FUNCTION_BLOCK Model (* Composite Function Block Type *)
  (* Standard: 61499-2 *)
  (* Version 0.0, 7/13/2016, Andrei, nxtControl GmbH, template *)
  PACKAGE Main;
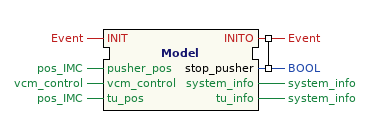
  EVENT_INPUT
    INIT; (* Initialization Request *)
  END_EVENT
  EVENT_OUTPUT
    INITO WITH stop_pusher; (* Initialization Confirm *)
  END_EVENT
  VAR_OUTPUT
    stop_pusher : BOOL;
  END_VAR
  SOCKETS
    pusher_pos : pos_IMC;
    vcm_control : vcm_control;
    tu_pos : pos_IMC;
  END_SOCKETS
  PLUGS
    system_info : system_info;
    tu_info : system_info;
  END_PLUGS
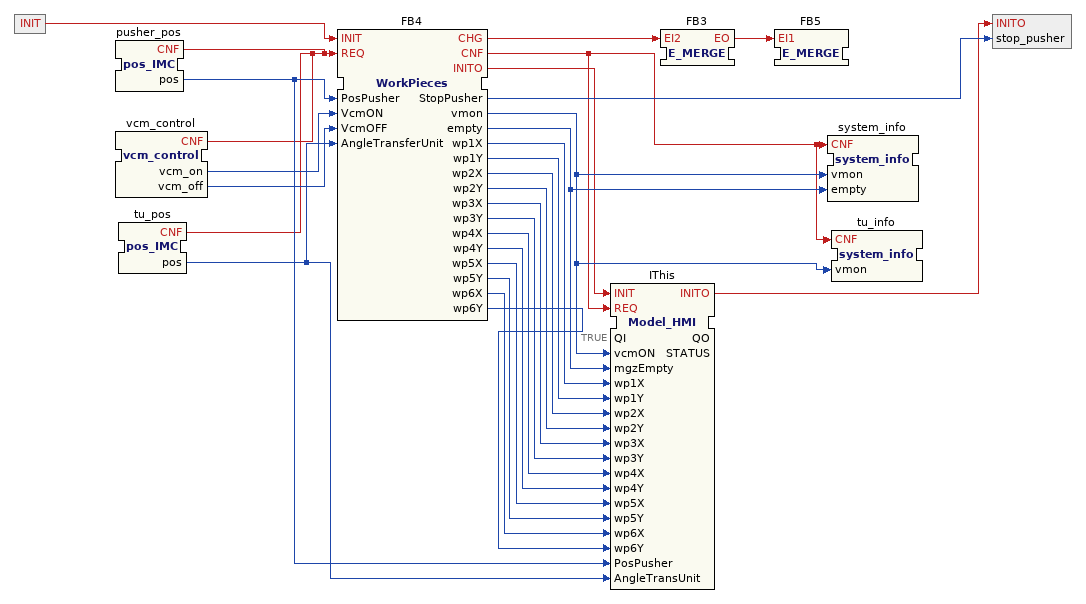
  FBS
    FB3 : E_MERGE;
    FB5 : E_MERGE;
    FB4 : WorkPieces;
    IThis : Model_HMI(QI := TRUE);
  END_FBS
  EVENT_CONNECTIONS
    FB4.CHG TO FB3.EI2;
    FB3.EO TO FB5.EI1;
    INIT TO FB4.INIT;
    pusher_pos.CNF TO FB4.REQ;
    vcm_control.CNF TO FB4.REQ;
    tu_pos.CNF TO FB4.REQ;
    FB4.CNF TO system_info.CNF;
    FB4.INITO TO IThis.INIT;
    FB4.CNF TO IThis.REQ;
    IThis.INITO TO INITO;
    FB4.CNF TO tu_info.CNF;
  END_CONNECTIONS
  DATA_CONNECTIONS
    FB4.StopPusher TO stop_pusher;
    pusher_pos.pos TO FB4.PosPusher;
    vcm_control.vcm_on TO FB4.VcmON;
    vcm_control.vcm_off TO FB4.VcmOFF;
    tu_pos.pos TO FB4.AngleTransferUnit;
    FB4.vmon TO system_info.vmon;
    FB4.empty TO system_info.empty;
    FB4.vmon TO IThis.vcmON;
    FB4.empty TO IThis.mgzEmpty;
    FB4.wp1X TO IThis.wp1X;
    FB4.wp1Y TO IThis.wp1Y;
    FB4.wp2X TO IThis.wp2X;
    FB4.wp2Y TO IThis.wp2Y;
    FB4.wp3X TO IThis.wp3X;
    FB4.wp3Y TO IThis.wp3Y;
    FB4.wp4X TO IThis.wp4X;
    FB4.wp4Y TO IThis.wp4Y;
    FB4.wp5X TO IThis.wp5X;
    FB4.wp5Y TO IThis.wp5Y;
    FB4.wp6X TO IThis.wp6X;
    FB4.wp6Y TO IThis.wp6Y;
    pusher_pos.pos TO IThis.PosPusher;
    tu_pos.pos TO IThis.AngleTransUnit;
    FB4.vmon TO tu_info.vmon;
  END_CONNECTIONS
END_FUNCTION_BLOCK
